SUBAPPLICATION Uebung_094d_AX (* OptionalGroup_001 OHNE DEMUX: die Gruppe ist immer aktiv, kein K/Index noetig - E_RESTART (COLD/WARM) loest einmalig INIT_REQ mit konstantem QI_OUT=TRUE aus, statt dass ein AOption_AUI_DEMUX_N je nach K einen von mehreren OUTx-Anschluessen waehlt. *)
  (* Standard: 61499-2; Description: Copyright (c) 2026 Meisterschulen am Ostbahnhof This program and the accompanying materials are made available under the terms of the Eclipse Public License 2.0 which is available at https://www.eclipse.org/legal/epl-2.0/ SPDX-License-Identifier: EPL-2.0 *)
  (* Version 1.0, 2026-10-15, Franz Höpfinger, Meisterschulen am Ostbahnhof, initial API and implementation and/or initial documentation *)
  PACKAGE Uebungen;
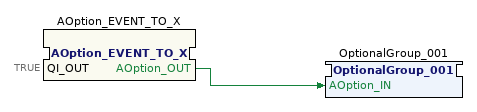
  FBS
    AOption_EVENT_TO_X : Option::conversion::AOption_EVENT_TO_X(QI_OUT := TRUE);
  END_FBS
  SUBAPPS
    OptionalGroup_001 : MyLib_AX_Option::sys::OptionalGroup_001;
  END_SUBAPPS
  ADAPTER_CONNECTIONS
    AOption_EVENT_TO_X.AOption_OUT TO OptionalGroup_001.AOption_IN;
  END_CONNECTIONS
END_SUBAPPLICATION
